SUBAPPLICATION mapping_aux (* Subapplication Type *)
  (* Standard: 61499-2 *)
  (* Version 1.0, 2023-01-29, Franz *)
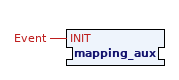
  EVENT_INPUT
    INIT;
  END_EVENT
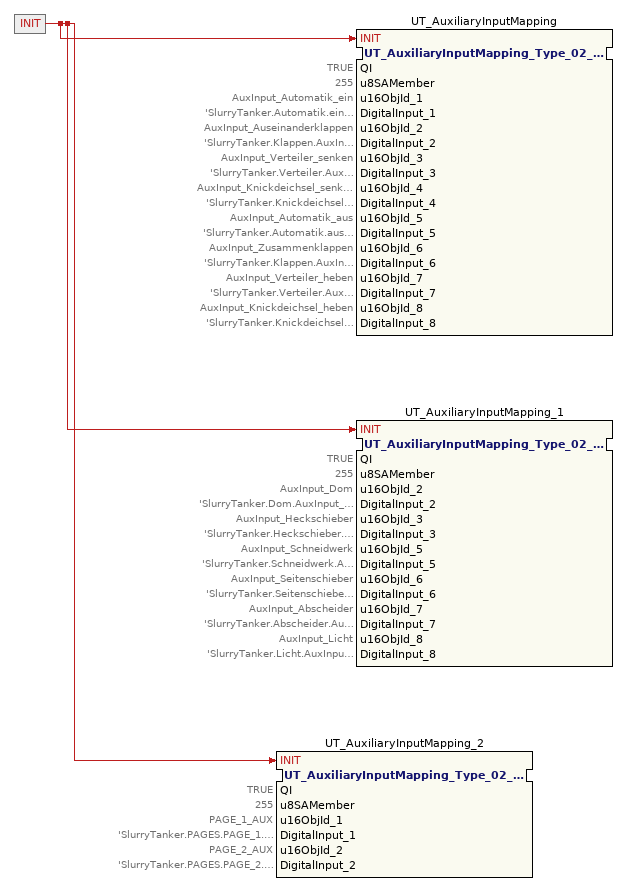
  FBS
    UT_AuxiliaryInputMapping : UT_AuxiliaryInputMapping_Type_02_Bool_NonLatched(QI := TRUE, u8SAMember := 255, u16ObjId_1 := AuxInput_Automatik_ein, DigitalInput_1 := 'SlurryTanker.Automatik.ein.AuxInput', u16ObjId_2 := AuxInput_Auseinanderklappen, DigitalInput_2 := 'SlurryTanker.Klappen.AuxInput_heben.AuxInput', u16ObjId_3 := AuxInput_Verteiler_senken, DigitalInput_3 := 'SlurryTanker.Verteiler.AuxInput_senken.AuxInput', u16ObjId_4 := AuxInput_Knickdeichsel_senken, DigitalInput_4 := 'SlurryTanker.Knickdeichsel.AuxInput_senken.AuxInput', u16ObjId_5 := AuxInput_Automatik_aus, DigitalInput_5 := 'SlurryTanker.Automatik.aus.AuxInput', u16ObjId_6 := AuxInput_Zusammenklappen, DigitalInput_6 := 'SlurryTanker.Klappen.AuxInput_senken.AuxInput', u16ObjId_7 := AuxInput_Verteiler_heben, DigitalInput_7 := 'SlurryTanker.Verteiler.AuxInput_heben.AuxInput', u16ObjId_8 := AuxInput_Knickdeichsel_heben, DigitalInput_8 := 'SlurryTanker.Knickdeichsel.AuxInput_heben.AuxInput');
    UT_AuxiliaryInputMapping_1 : UT_AuxiliaryInputMapping_Type_02_Bool_NonLatched(QI := TRUE, u8SAMember := 255, u16ObjId_2 := AuxInput_Dom, DigitalInput_2 := 'SlurryTanker.Dom.AuxInput_UP.AuxInput', u16ObjId_3 := AuxInput_Heckschieber, DigitalInput_3 := 'SlurryTanker.Heckschieber.AuxInput_UP.AuxInput', u16ObjId_5 := AuxInput_Schneidwerk, DigitalInput_5 := 'SlurryTanker.Schneidwerk.AuxInput_UP.AuxInput', u16ObjId_6 := AuxInput_Seitenschieber, DigitalInput_6 := 'SlurryTanker.Seitenschieber.AuxInput_UP.AuxInput', u16ObjId_7 := AuxInput_Abscheider, DigitalInput_7 := 'SlurryTanker.Abscheider.AuxInput_UP.AuxInput', u16ObjId_8 := AuxInput_Licht, DigitalInput_8 := 'SlurryTanker.Licht.AuxInput_UP.AuxInput');
    UT_AuxiliaryInputMapping_2 : UT_AuxiliaryInputMapping_Type_02_Bool_NonLatched(QI := TRUE, u8SAMember := 255, u16ObjId_1 := PAGE_1_AUX, DigitalInput_1 := 'SlurryTanker.PAGES.PAGE_1.AUX', u16ObjId_2 := PAGE_2_AUX, DigitalInput_2 := 'SlurryTanker.PAGES.PAGE_2.AUX');
  END_FBS
  EVENT_CONNECTIONS
    INIT TO UT_AuxiliaryInputMapping.INIT;
    INIT TO UT_AuxiliaryInputMapping_1.INIT;
    INIT TO UT_AuxiliaryInputMapping_2.INIT;
  END_CONNECTIONS
END_SUBAPPLICATION
